TYPE ST_LightCommand :
STRUCT
    bValid : BOOL;
    bOn : BOOL;
END_STRUCT
END_TYPE

(* stored: Version 1.1.0.1
   DUT ST_LightCommand: Id {60bcb23a-88c4-4222-baa8-3b0937aa8ff1} *)
